(* IEC 61131-3 sources: llm-plc-st-eval/data/definitivo/gemini-3.1-pro-preview/B6/zero_shot, 3 files *)

(* ---- ejec_1.st ---- *)
```iecst
FUNCTION_BLOCK FB_Baliza
VAR_INPUT
    alarma : BOOL; // Condición de alarma activa
END_VAR
VAR_OUTPUT
    lampara : BOOL; // Salida hacia la baliza luminosa
END_VAR
VAR
    Timer_ON : TON; // Temporizador para el tiempo de encendido (1s)
    Timer_OFF : TON; // Temporizador para el tiempo de apagado (1s)
END_VAR

// Temporizador que cuenta el tiempo que la lámpara permanece encendida
Timer_ON(IN := alarma AND NOT Timer_OFF.Q, PT := T#1S);

// Temporizador que cuenta el tiempo que la lámpara permanece apagada
Timer_OFF(IN := Timer_ON.Q, PT := T#1S);

// La lámpara enciende inmediatamente con la alarma y alterna su estado cada segundo
lampara := alarma AND NOT Timer_ON.Q;

END_FUNCTION_BLOCK
```

(* ---- ejec_2.st ---- *)
```iecst
FUNCTION_BLOCK FB_Baliza
VAR_INPUT
    alarma : BOOL; (* Condición de activación de la alarma *)
END_VAR
VAR_OUTPUT
    lampara : BOOL; (* Estado de la baliza luminosa *)
END_VAR
VAR
    tonEncendido : TON; (* Temporizador para el ciclo de encendido *)
    tonApagado : TON;   (* Temporizador para el ciclo de apagado *)
END_VAR

(* El primer temporizador cuenta 1s mientras la alarma esté activa y el segundo no haya terminado *)
tonEncendido(IN := alarma AND NOT tonApagado.Q, PT := T#1S);

(* El segundo temporizador cuenta 1s después de que el primero termina *)
tonApagado(IN := tonEncendido.Q, PT := T#1S);

(* La lámpara se enciende inmediatamente con la alarma y se apaga al terminar el primer tiempo *)
lampara := alarma AND NOT tonEncendido.Q;

END_FUNCTION_BLOCK
```

(* ---- ejec_3.st ---- *)
```iecst
FUNCTION_BLOCK FB_Baliza
VAR_INPUT
    alarma : BOOL; // Condicion de activacion de la alarma
END_VAR
VAR_OUTPUT
    lampara : BOOL; // Salida hacia la baliza luminosa
END_VAR
VAR
    ton_Encendido : TON; // Temporizador para el tiempo en estado encendido
    ton_Apagado : TON;   // Temporizador para el tiempo en estado apagado
END_VAR

// Generador de ciclo: ton_Encendido se activa con la alarma y se reinicia con ton_Apagado
ton_Encendido(IN := alarma AND NOT ton_Apagado.Q, PT := T#1S);

// ton_Apagado comienza a contar cuando ton_Encendido alcanza 1 segundo
ton_Apagado(IN := ton_Encendido.Q, PT := T#1S);

// La lampara se enciende si hay alarma, y se apaga durante el ciclo de ton_Apagado
lampara := alarma AND NOT ton_Encendido.Q;

END_FUNCTION_BLOCK
```
